(* CODESYS project snapshot.xml
   cds-daemon-config: {"poll_ms": 60, "deny": []}
   cts-project-id: 374e2afd-b7d6-4447-8bd8-ce8e480d827d
   cds-sync-pc: WIN-CODESYS
   cds-sync-folder: ..

Project tree, tasks and I/O mapping:
  PLC_Stabur : PLC Stabur, PSV Electric, order no. psve.ru, version 3.5.16.40
    application Application
      libraries: SysTimeCore, * (System); CmpLog, * (System); CmpErrors, * (System); CmpApp, * (System); Standard, 3.5.22.0 (System); Component Manager, * (System); CmpIecTask, * (System)
      task VISU_TASK (cyclic, interval 100 ms, priority 31) calls VisuElems.Visu_Prg
      task Task (cyclic, interval 200 ms, priority 1) calls MAIN
      data type ST_Bits8
      data type ST_Packed
      function block FB_Logger [ST]: LogADDLong, LogSafe, LogADD, Fmt100
      data type U_Bits8
      program PRG_BitBench [ST]
      visualisation Visualization
      global variables LogComponent
      program MAIN [ST]
      function block FB_BenchRun [ST]
      data type ST_Bools8
      global variables GVL_Bench
      data type U_ExtBits
      data type ST_Bits8Ext
      data type E_BenchMode
      function block FB_Motor [ST]
      global variables GVL_Motors
      function F_Scale [ST]
      global variables GVL_Fixture
      function block FB_Valve [ST]: P_Open, A_Reset, M_Toggle
      LiveTmpFolder/
        global variables GVL_LiveTmp
      interface I_LiveTmp: M_LiveTmp
    Retain_ : Retain, PSV Electric, order no. --0--, version 3.5.16.40
        unmapped channels: Record counter, RETAIN status code, Write
    Leds : Leds, PSV Electro, order no. --0--, version 3.5.16.40
        unmapped channels: LEDs, Screen brightness, Buzzer
  text list GlobalTextList
*)

// PLC_Stabur/Application/ST_Bits8
TYPE ST_Bits8 :
STRUCT
	bit0 : BIT;
	bit1 : BIT;
	bit2 : BIT;
	bit3 : BIT;
	bit4 : BIT;
	bit5 : BIT;
	bit6 : BIT;
	bit7 : BIT;
END_STRUCT
END_TYPE

// PLC_Stabur/Application/ST_Packed
{attribute 'pack_mode' := '0'}
TYPE ST_Packed :
STRUCT
	bTag : BOOL;
	wData : WORD;
END_STRUCT
END_TYPE

// PLC_Stabur/Application/U_Bits8
TYPE U_Bits8 :
UNION
	b : BYTE;
	bits : ST_Bits8;
END_UNION
END_TYPE

// PLC_Stabur/Application/ST_Bools8
TYPE ST_Bools8 :
STRUCT
	b0 : BOOL;
	b1 : BOOL;
	b2 : BOOL;
	b3 : BOOL;
	b4 : BOOL;
	b5 : BOOL;
	b6 : BOOL;
	b7 : BOOL;
END_STRUCT
END_TYPE

// PLC_Stabur/Application/U_ExtBits
TYPE U_ExtBits :
UNION
	b : BYTE;
	bits : ST_Bits8Ext;
END_UNION
END_TYPE

// PLC_Stabur/Application/ST_Bits8Ext
TYPE ST_Bits8Ext EXTENDS ST_Bits8 :
STRUCT
END_STRUCT
END_TYPE

// PLC_Stabur/Application/E_BenchMode
{attribute 'qualified_only'}
TYPE E_BenchMode :
(
	Idle := 0,
	Run := 1,
	Fault := 7
) INT;
END_TYPE

// PLC_Stabur/Application/LogComponent
{attribute 'qualified_only'}
{attribute 'symbol' := 'none'}
VAR_GLOBAL
	BITBENCH : STRING := 'BitBench';	// component name in the runtime log
	sNumFmt  : STRING(80);				// FB_Logger.Fmt100 puts the formatted number here

	logger : FB_Logger;					// the logger itself (production sample)
END_VAR

// PLC_Stabur/Application/GVL_Bench
{attribute 'qualified_only'}
VAR_GLOBAL
	// --- control (written by the host; a run starts itself 50 cycles after start) ---
	xRun			: BOOL;			// rising edge: run the tests again
	xRunUnaligned	: BOOL;			// TRUE: also run B8 (unaligned WORD, may crash)
	sCpuMode		: STRING(40);	// CPU frequency mode, written by the host before a run; printed in the log
	// --- observation ---
	xDone			: BOOL;			// run finished
	nState			: INT;			// state of the PRG_BitBench machine
	nTestIdx		: INT;			// current test 0..21 (a round = one test in one cycle)
	nMeasIdx		: INT;			// how many pairs went into the statistics of the last round
	nIter			: UDINT;		// iterations in one half of a pair (both halves are identical)
	nHeartbeat		: UDINT;		// ++ on every call of the task
	nLastNs			: ULINT;		// duration of the last round (without calibration), ns
	dwSink			: DWORD;		// read sink
	dwSinkW			: DWORD;		// write sink (write baseline)
	// --- results: index 0..10 = B0..B7c, B8 ---
	// Difference = variant - base within a pair, the unit is HUNDREDTHS of ns/operation.
	// The median and the percentiles are computed over the pair differences of one round (NPAIRS = 101).
	medDiffRead		: ARRAY [0..10] OF DINT;	// median of the difference, read
	p25DiffRead		: ARRAY [0..10] OF DINT;	// 25th percentile of the difference
	p75DiffRead		: ARRAY [0..10] OF DINT;	// 75th percentile of the difference
	minDiffRead		: ARRAY [0..10] OF DINT;	// the smallest difference (extreme point)
	minVarRead		: ARRAY [0..10] OF DWORD;	// absolute minimum of the variant, hundredths of ns/op
	minBaseRead		: ARRAY [0..10] OF DWORD;	// absolute minimum of the base, hundredths of ns/op
	nIterRead		: ARRAY [0..10] OF UDINT;	// nIter at the end of the test
	nRoundUsRead	: ARRAY [0..10] OF UDINT;	// duration of the round, us
	medDiffWrite	: ARRAY [0..10] OF DINT;	// median of the difference, write
	p25DiffWrite	: ARRAY [0..10] OF DINT;
	p75DiffWrite	: ARRAY [0..10] OF DINT;
	minDiffWrite	: ARRAY [0..10] OF DINT;
	minVarWrite		: ARRAY [0..10] OF DWORD;
	minBaseWrite	: ARRAY [0..10] OF DWORD;
	nIterWrite		: ARRAY [0..10] OF UDINT;
	nRoundUsWrite	: ARRAY [0..10] OF UDINT;
	nMeasDone		: ARRAY [0..10] OF INT;		// how many pairs went into the result (0 = SKIPPED)
	// --- one-off values ---
	aSizeof			: ARRAY [0..5] OF INT;		// SIZEOF of the types
	// --- enum live check ---
	eMode : E_BenchMode := E_BenchMode.Idle;
	aMode : ARRAY [0..2] OF E_BenchMode := [E_BenchMode.Idle, E_BenchMode.Run, E_BenchMode.Fault];
	// --- test data ---
	stBools			: ST_Bools8;
	stBits			: ST_Bits8;
	uBits			: U_Bits8;
	uExt			: U_ExtBits;
	wData			: WORD;
	dwDataB6		: DWORD;
	stPacked		: ST_Packed;
END_VAR

// PLC_Stabur/Application/GVL_Motors
{attribute 'qualified_only'}
VAR_GLOBAL
	xM1Start : BOOL;
	xM1Stop : BOOL;
	xM1Feedback : BOOL;
	xM1Reset : BOOL;
	xM1Run : BOOL;
	xM1Fault : BOOL;
	nM1Starts : UDINT;
	fbMotor1 : FB_Motor;

	xM2Start : BOOL;
	xM2Stop : BOOL;
	xM2Feedback : BOOL;
	xM2Reset : BOOL;
	xM2Run : BOOL;
	xM2Fault : BOOL;
	nM2Starts : UDINT;
	fbMotor2 : FB_Motor;
END_VAR

// PLC_Stabur/Application/GVL_Fixture
VAR_GLOBAL
	rScaled : REAL;
	xValveOpen : BOOL;
	fbValve : FB_Valve;
	nTicks : UDINT;
END_VAR

// PLC_Stabur/Application/LiveTmpFolder/GVL_LiveTmp
VAR_GLOBAL
	xLiveTmp : BOOL;
END_VAR

// PLC_Stabur/Application/MAIN
PROGRAM MAIN
(* t76 timing probe *)
VAR
	eObservedMode : E_BenchMode;
END_VAR

// Self-contained bit-access benchmark: it starts itself 50 cycles after the
// application starts, writes its report to the runtime log, and repeats on GVL_Bench.xRun.
// Project created with the cds-text-sync daemon and LLM agent.
PRG_BitBench();
eObservedMode := GVL_Bench.eMode;

GVL_Motors.fbMotor1(
	xStart := GVL_Motors.xM1Start,
	xStop := GVL_Motors.xM1Stop,
	xFeedback := GVL_Motors.xM1Feedback,
	xReset := GVL_Motors.xM1Reset,
	xRun => GVL_Motors.xM1Run,
	xFault => GVL_Motors.xM1Fault,
	nStarts => GVL_Motors.nM1Starts);
GVL_Motors.fbMotor2(
	xStart := GVL_Motors.xM2Start,
	xStop := GVL_Motors.xM2Stop,
	xFeedback := GVL_Motors.xM2Feedback,
	xReset := GVL_Motors.xM2Reset,
	xRun => GVL_Motors.xM2Run,
	xFault => GVL_Motors.xM2Fault,
	nStarts => GVL_Motors.nM2Starts);

// Fixture: exercise the function, property, action and interface kinds.
GVL_Fixture.nTicks := GVL_Fixture.nTicks + 1;
GVL_Fixture.rScaled := F_Scale(UDINT_TO_REAL(GVL_Fixture.nTicks), 0.5);
IF GVL_Fixture.nTicks MOD 10 = 0 THEN
	GVL_Fixture.fbValve.M_Toggle();
END_IF
GVL_Fixture.xValveOpen := GVL_Fixture.fbValve.P_Open;

END_PROGRAM

// PLC_Stabur/Application/PRG_BitBench
(*
BitBench — a self-contained benchmark of the cost of bit access.

Project created with the cds-text-sync daemon and LLM agent.
Bench: PLC_Stabur (RK3568, 4x ARM Cortex-A55), CODESYS Control 3.5.16.40,
task t#200 ms, timer SysTimeGetNs on the PLC.

RUN ORDER (counted in task cycles):
  PLC on / application started
  -> wait START_WAIT cycles (50 = 10 s)
  -> round 1: one test ENTIRELY in one cycle
  -> wait GAP_WAIT cycles (5 = 1 s)
  -> round 2 ... and so on up to the last test
  -> conclusion (Conclusion) and 'BitBench: done'.
The 20 tests (B0..B7c read and write) take about 30 s; B8 takes two more rounds.

THE METHOD OF ONE ROUND - PAIRED MEASUREMENTS.
The calibration (CAL_N iterations) chooses nIter so that one half of a pair runs
for about TARGET_EACH_NS. Then WARM_PAIRS warm-up pairs and NPAIRS measured pairs
in a row: a pair is the baseline and the variant with the same nIter, the order
alternates (even pair base -> variant, odd pair the other way round). The result
of a pair is the difference (variant - base) in hundredths of ns/operation. The
differences are sorted at the end of the round; Result is the median, with p25,
p75 and min beside it.

A round is limited by ROUND_BUDGET_NS: if the pairs did not fit, the round is cut
short and is computed from the pairs that made it (fewer than MIN_PAIRS -
SKIPPED). We reset the statistics of the task (CmpIecTask) in the last cycle of
the pause before the round and read them in the first cycle after it: the cycle
max is the round itself.

Restart. A run starts over (from the START_WAIT pause) if:
  - the application was downloaded or reset (the variables are initialised);
  - more than RESTART_GAP_NS passed between two cycles (Online -> Stop/Start:
    the variables survive, but the task was stopped);
  - a rising edge on GVL_Bench.xRun (then the pause is GAP_WAIT, not START_WAIT).
B8 (an unaligned WORD in a STRUCT with pack_mode 0) runs only when
GVL_Bench.xRunUnaligned is set, because it may raise an exception.

We keep the log strings no longer than 120 characters (the runtime cuts a record
at 127); anything longer is sent by LogSafe in pieces.
*)

PROGRAM PRG_BitBench
VAR CONSTANT
	// --- schedule, in task cycles ---
	START_WAIT	: INT := 50;			// after the application starts
	GAP_WAIT	: INT := 5;				// between rounds
	TASK_NS		: ULINT := 200000000;	// task period, ns (t#200 ms)
	RESTART_GAP_NS : ULINT := 1000000000;	// a gap between cycles longer than 1 s = the task was stopped
	// --- method ---
	CAL_N		: UDINT := 1000;		// iterations in the calibration half
	WARM_PAIRS	: INT := 5;				// warm-up pairs (they do not enter the statistics)
	NPAIRS		: INT := 101;			// measured pairs per test (odd - the median is unambiguous)
	MIN_PAIRS	: INT := 21;			// fewer - the test is SKIPPED
	MIN_ITER	: UDINT := 50;
	MAX_ITER	: UDINT := 2000000;
	TARGET_EACH_NS : ULINT := 200000;	// target duration of half a pair, ns (0.2 ms)
	ROUND_BUDGET_NS : ULINT := 80000000;	// round limit, ns (80 ms = 40 % of the cycle)
	// --- tests ---
	IDX_LAST_MAIN : INT := 19;			// 0..9 read B0..B7c, 10..19 write
	IDX_LAST	: INT := 21;			// 20 = read B8, 21 = write B8
	// --- states ---
	ST_IDLE		: INT := 0;				// no run in progress
	ST_WAIT		: INT := 10;			// pause before a round (nWait cycles)
	ST_ROUND	: INT := 20;			// round: one test in this cycle
	ST_DONE		: INT := 100;			// run finished
END_VAR
VAR
	// --- start and restart ---
	xInit		: BOOL;			// FALSE after a download/reset: the first cycle
	xRunPrev	: BOOL;
	tNow		: ULINT;
	tPrevCycle	: ULINT;
	// --- state machine ---
	nFsm		: INT;
	nWait		: INT;			// how many cycles of the pause are left
	xHeadDone	: BOOL;			// the run header has already been printed
	xStatPending : BOOL;		// print the statistics of the task for the round in this cycle
	nTestNo		: INT;			// 0..21
	// --- current test ---
	nMode		: INT;			// 0 = read, 1 = write
	nVariant	: INT;			// 0..10
	nIterCur	: UDINT;		// nIter of the round: the same for both halves of every pair
	// --- statistics of the task itself (CmpIecTask, as in FB_TaskInfo from a production sample) ---
	pTaskInfo	: POINTER TO Task_Info2;
	resTask		: UDINT;
	// --- measurements ---
	fbRun		: FB_BenchRun;
	tBase		: ULINT;
	tVar		: ULINT;
	tPair		: ULINT;
	tRound0		: ULINT;
	tRoundNs	: ULINT;		// duration of the round (without calibration), ns
	uCalBase	: ULINT;
	uCalVar		: ULINT;
	aDiff		: ARRAY [0..100] OF DINT;	// pair differences (NPAIRS = 101)
	nMeasCnt	: INT;
	xCut		: BOOL;			// the round was cut by ROUND_BUDGET_NS
	uMaxPair	: ULINT;
	uMinVar		: ULINT;		// absolute minimum of the variant, hundredths of ns/op
	uMinBase	: ULINT;
	dNew		: DINT;
	dMed		: DINT;
	dP25		: DINT;
	dP75		: DINT;
	dMn			: DINT;
	// --- processing ---
	p			: INT;
	i			: INT;
	j			: INT;
	uTmp		: ULINT;
	dwRes		: DWORD;
	xTimerBad	: BOOL;
	dRead		: DINT;
	dWrite		: DINT;
	dWorst		: DINT;
	dTmp		: DINT;
	// --- strings ---
	sMsg		: STRING(255);
	sName		: STRING(40);
	sWhat		: STRING(80);
END_VAR

// ===================== 1. start, restart, manual run =====================
dwRes := SysTimeGetNs(tNow);

IF NOT xInit THEN
	// the first cycle after a download or a reset
	xInit := TRUE;
	nFsm := ST_WAIT;
	nWait := START_WAIT;
	xHeadDone := FALSE;
	xStatPending := FALSE;
	LogComponent.logger.LogSafe(LogComponent.BITBENCH, CmpLog.LogClass.LOG_INFO,
		'BitBench: application started, first round after 50 cycles');
ELSIF tPrevCycle <> 0 AND tNow - tPrevCycle > RESTART_GAP_NS THEN
	// the task was stopped (Online -> Stop/Start): we start the run over
	nFsm := ST_WAIT;
	nWait := START_WAIT;
	xHeadDone := FALSE;
	xStatPending := FALSE;
	LogComponent.logger.LogSafe(LogComponent.BITBENCH, CmpLog.LogClass.LOG_INFO,
		'BitBench: restart after a stop, first round after 50 cycles');
END_IF
tPrevCycle := tNow;

IF GVL_Bench.xRun AND NOT xRunPrev THEN
	nFsm := ST_WAIT;
	nWait := GAP_WAIT;
	xHeadDone := FALSE;
	xStatPending := FALSE;
END_IF
xRunPrev := GVL_Bench.xRun;

// ===================== 2. task statistics for the previous round =====================
IF xStatPending THEN
	xStatPending := FALSE;
	IF pTaskInfo <> 0 THEN
		sMsg := CONCAT('Task      ', sName);
		sMsg := CONCAT(sMsg, ': cycle max ');
		sMsg := CONCAT(sMsg, DWORD_TO_STRING(pTaskInfo^.dwMaxCycleTime));
		sMsg := CONCAT(sMsg, ' us, jitter max ');
		sMsg := CONCAT(sMsg, DINT_TO_STRING(pTaskInfo^.iJitterMax));
		sMsg := CONCAT(sMsg, ' us, min ');
		sMsg := CONCAT(sMsg, DINT_TO_STRING(pTaskInfo^.iJitterMin));
		sMsg := CONCAT(sMsg, ' us');
		LogComponent.logger.LogSafe(LogComponent.BITBENCH, CmpLog.LogClass.LOG_INFO, sMsg);
	END_IF
END_IF

// ===================== 3. state machine =====================
CASE nFsm OF
ST_IDLE:
	;	// waiting for xRun or a restart

ST_WAIT:	// pause; the last cycle of the pause prepares the round
	nWait := nWait - 1;
	IF nWait <= 0 THEN
		IF NOT xHeadDone THEN
			xHeadDone := TRUE;
			nTestNo := 0;
			xTimerBad := FALSE;
			GVL_Bench.xDone := FALSE;
			GVL_Bench.dwSink := 0;
			GVL_Bench.dwSinkW := 0;
			// clear the results of the previous run: after a SKIPPED or a crash
			// the GVL must not keep numbers from the previous run
			FOR i := 0 TO 10 DO
				GVL_Bench.medDiffRead[i] := 0;
				GVL_Bench.p25DiffRead[i] := 0;
				GVL_Bench.p75DiffRead[i] := 0;
				GVL_Bench.minDiffRead[i] := 0;
				GVL_Bench.minVarRead[i] := 0;
				GVL_Bench.minBaseRead[i] := 0;
				GVL_Bench.nIterRead[i] := 0;
				GVL_Bench.nRoundUsRead[i] := 0;
				GVL_Bench.medDiffWrite[i] := 0;
				GVL_Bench.p25DiffWrite[i] := 0;
				GVL_Bench.p75DiffWrite[i] := 0;
				GVL_Bench.minDiffWrite[i] := 0;
				GVL_Bench.minVarWrite[i] := 0;
				GVL_Bench.minBaseWrite[i] := 0;
				GVL_Bench.nIterWrite[i] := 0;
				GVL_Bench.nRoundUsWrite[i] := 0;
				GVL_Bench.nMeasDone[i] := 0;
			END_FOR
			GVL_Bench.nIter := 0;
			GVL_Bench.nLastNs := 0;
			GVL_Bench.nMeasIdx := 0;

			// the run header
			LogComponent.logger.LogSafe(LogComponent.BITBENCH, CmpLog.LogClass.LOG_INFO,
				'BitBench: project created with cds-text-sync daemon and LLM agent');

			sMsg := CONCAT('BitBench: start, CPU mode ', GVL_Bench.sCpuMode);
			LogComponent.logger.LogSafe(LogComponent.BITBENCH, CmpLog.LogClass.LOG_INFO, sMsg);

			sMsg := 'BitBench: CPU RK3568 4x ARM Cortex-A55, task t#';
			sMsg := CONCAT(sMsg, ULINT_TO_STRING(TASK_NS / 1000000));
			sMsg := CONCAT(sMsg, ' ms, timer SysTimeGetNs on the PLC');
			LogComponent.logger.LogSafe(LogComponent.BITBENCH, CmpLog.LogClass.LOG_INFO, sMsg);

			sMsg := 'BitBench: 1 round = 1 test in one cycle, ';
			sMsg := CONCAT(sMsg, INT_TO_STRING(GAP_WAIT));
			sMsg := CONCAT(sMsg, ' cycles between rounds, round limit ');
			sMsg := CONCAT(sMsg, ULINT_TO_STRING(ROUND_BUDGET_NS / 1000000));
			sMsg := CONCAT(sMsg, ' ms');
			LogComponent.logger.LogSafe(LogComponent.BITBENCH, CmpLog.LogClass.LOG_INFO, sMsg);

			sMsg := 'BitBench: round = ';
			sMsg := CONCAT(sMsg, INT_TO_STRING(WARM_PAIRS));
			sMsg := CONCAT(sMsg, ' warm-up + ');
			sMsg := CONCAT(sMsg, INT_TO_STRING(NPAIRS));
			sMsg := CONCAT(sMsg, ' measured pairs (base and variant, same nIter), half ~');
			LogComponent.logger.Fmt100(ULINT_TO_DINT(TARGET_EACH_NS / 10000), FALSE);
			sMsg := CONCAT(sMsg, LogComponent.sNumFmt);
			sMsg := CONCAT(sMsg, ' ms');
			LogComponent.logger.LogSafe(LogComponent.BITBENCH, CmpLog.LogClass.LOG_INFO, sMsg);

			GVL_Bench.aSizeof[0] := SIZEOF(GVL_Bench.stBools);
			GVL_Bench.aSizeof[1] := SIZEOF(GVL_Bench.stBits);
			GVL_Bench.aSizeof[2] := SIZEOF(GVL_Bench.uBits);
			GVL_Bench.aSizeof[3] := SIZEOF(GVL_Bench.uExt);
			GVL_Bench.aSizeof[4] := SIZEOF(GVL_Bench.stPacked);
			GVL_Bench.aSizeof[5] := SIZEOF(GVL_Bench.wData);

			sMsg := 'Memory: 8 BOOL in a STRUCT = ';
			sMsg := CONCAT(sMsg, INT_TO_STRING(GVL_Bench.aSizeof[0]));
			sMsg := CONCAT(sMsg, ' B, 8 BIT in a STRUCT = ');
			sMsg := CONCAT(sMsg, INT_TO_STRING(GVL_Bench.aSizeof[1]));
			sMsg := CONCAT(sMsg, ' B, UNION of 8 BIT = ');
			sMsg := CONCAT(sMsg, INT_TO_STRING(GVL_Bench.aSizeof[2]));
			sMsg := CONCAT(sMsg, ' B');
			LogComponent.logger.LogSafe(LogComponent.BITBENCH, CmpLog.LogClass.LOG_INFO, sMsg);

			sMsg := 'Memory: the same UNION + EXTENDS = ';
			sMsg := CONCAT(sMsg, INT_TO_STRING(GVL_Bench.aSizeof[3]));
			sMsg := CONCAT(sMsg, ' B, WORD = ');
			sMsg := CONCAT(sMsg, INT_TO_STRING(GVL_Bench.aSizeof[5]));
			sMsg := CONCAT(sMsg, ' B, pack_mode 0 (WORD after BOOL) = ');
			sMsg := CONCAT(sMsg, INT_TO_STRING(GVL_Bench.aSizeof[4]));
			sMsg := CONCAT(sMsg, ' B');
			LogComponent.logger.LogSafe(LogComponent.BITBENCH, CmpLog.LogClass.LOG_INFO, sMsg);

			LogComponent.logger.LogSafe(LogComponent.BITBENCH, CmpLog.LogClass.LOG_INFO,
				'Base  read: dwSink := dwSink + 1; write: dwSinkW := UDINT_TO_DWORD(k AND 1)');

			IF pTaskInfo = 0 THEN
				pTaskInfo := IecTaskGetInfo3(hIecTask := IecTaskGetCurrent(ADR(resTask)),
				                             pResult := ADR(resTask));
			END_IF
		END_IF

		// the task statistics from this moment on are the statistics of the round
		IecTaskResetStatistics(IecTaskGetCurrent(ADR(resTask)));
		nFsm := ST_ROUND;
	END_IF

ST_ROUND:	// one test entirely in this cycle
	// ---------- which test ----------
	IF nTestNo < 10 THEN
		nMode := 0;
		nVariant := nTestNo;
	ELSIF nTestNo <= IDX_LAST_MAIN THEN
		nMode := 1;
		nVariant := nTestNo - 10;
	ELSIF nTestNo = IDX_LAST_MAIN + 1 THEN
		nMode := 0;
		nVariant := 10;
	ELSE
		nMode := 1;
		nVariant := 10;
	END_IF

	CASE nVariant OF
	0:	sName := 'B0 empty loop';
		sWhat := 'control: the variant is the base itself, expect 0';
	1:	sName := 'B1 BOOL fields';
		sWhat := '8 BOOL in a STRUCT, 1 byte each - the reference for the bit tests';
	2:	sName := 'B2 BIT fields';
		sWhat := '8 BIT packed into 1 byte - the write is a read-modify-write';
	3:	sName := 'B3 UNION+EXTENDS';
		sWhat := 'bit via a UNION that EXTENDS ST_Bits8; watch C0542';
	4:	sName := 'B4 UNION';
		sWhat := 'the same 8 BIT in a UNION, without EXTENDS';
	5:	sName := 'B5 WORD.3';
		sWhat := 'bit access to a WORD by dot: wData.3, 16 bits in 2 B';
	6:	sName := 'B6 mask var index';
		sWhat := 'mask (SHR(dwData, i) AND 1), no bit instruction';
	7:	sName := 'B7a 8 BOOL';
		sWhat := '8 BOOL one by one - one iteration = 8 accesses';
	8:	sName := 'B7b byte';
		sWhat := 'all 8 bits as one BYTE - one iteration = 1 access';
	9:	sName := 'B7c word';
		sWhat := 'all 16 bits as one WORD - one iteration = 1 access';
	10:	sName := 'B8 unaligned WORD';
		sWhat := 'pack_mode 0, wData.3 unaligned - the test may raise an exception';
	ELSE
		sName := 'B? unknown';
		sWhat := 'unknown variant';
	END_CASE

	sMsg := CONCAT('Testing ', sName);
	IF nMode = 0 THEN
		sMsg := CONCAT(sMsg, ' (read): ');
	ELSE
		sMsg := CONCAT(sMsg, ' (write): ');
	END_IF
	sMsg := CONCAT(sMsg, sWhat);
	LogComponent.logger.LogSafe(LogComponent.BITBENCH, CmpLog.LogClass.LOG_INFO, sMsg);

	IF nVariant = 10 THEN
		LogComponent.logger.LogSafe(LogComponent.BITBENCH, CmpLog.LogClass.LOG_WARNING,
			'B8 warning: unaligned WORD in a STRUCT with pack_mode 0; an exception here means the app restarts');
	END_IF

	// ---------- calibration: nIter for TARGET_EACH_NS from the slower half ----------
	fbRun(nWhich := 0, nMode := nMode, nVariant := nVariant, nIter := CAL_N);
	uCalBase := fbRun.tDur;
	IF fbRun.dwRes <> 0 THEN
		dwRes := fbRun.dwRes;
	END_IF
	fbRun(nWhich := 1, nMode := nMode, nVariant := nVariant, nIter := CAL_N);
	uCalVar := fbRun.tDur;
	IF fbRun.dwRes <> 0 THEN
		dwRes := fbRun.dwRes;
	END_IF

	uTmp := uCalBase;
	IF uCalVar > uTmp THEN
		uTmp := uCalVar;
	END_IF
	IF uTmp <> 0 THEN
		uTmp := (TARGET_EACH_NS * CAL_N) / uTmp;
	ELSE
		uTmp := MIN_ITER;
	END_IF
	IF uTmp < MIN_ITER THEN
		uTmp := MIN_ITER;
	END_IF
	IF uTmp > MAX_ITER THEN
		uTmp := MAX_ITER;
	END_IF
	nIterCur := ULINT_TO_UDINT(uTmp);
	GVL_Bench.nIter := nIterCur;

	// ---------- pairs: warm-up, then measured ----------
	nMeasCnt := 0;
	xCut := FALSE;
	uMaxPair := 0;
	uMinVar := 16#FFFFFFFFFFFFFFFF;
	uMinBase := 16#FFFFFFFFFFFFFFFF;
	SysTimeGetNs(tRound0);

	FOR p := 0 TO WARM_PAIRS + NPAIRS - 1 DO
		IF (p MOD 2) = 0 THEN
			fbRun(nWhich := 0, nMode := nMode, nVariant := nVariant, nIter := nIterCur);
			tBase := fbRun.tDur;
			fbRun(nWhich := 1, nMode := nMode, nVariant := nVariant, nIter := nIterCur);
			tVar := fbRun.tDur;
		ELSE
			fbRun(nWhich := 1, nMode := nMode, nVariant := nVariant, nIter := nIterCur);
			tVar := fbRun.tDur;
			fbRun(nWhich := 0, nMode := nMode, nVariant := nVariant, nIter := nIterCur);
			tBase := fbRun.tDur;
		END_IF
		IF fbRun.dwRes <> 0 THEN
			dwRes := fbRun.dwRes;
		END_IF

		IF p >= WARM_PAIRS THEN
			tPair := tBase + tVar;
			IF tPair > uMaxPair THEN
				uMaxPair := tPair;
			END_IF
			// the difference in hundredths of ns/op: each half is normalised separately
			uTmp := (tVar * 100) / nIterCur;
			IF uTmp < uMinVar THEN
				uMinVar := uTmp;
			END_IF
			dNew := ULINT_TO_DINT(uTmp);
			uTmp := (tBase * 100) / nIterCur;
			IF uTmp < uMinBase THEN
				uMinBase := uTmp;
			END_IF
			dNew := dNew - ULINT_TO_DINT(uTmp);
			aDiff[nMeasCnt] := dNew;
			nMeasCnt := nMeasCnt + 1;
		END_IF

		// round limit: the task cycle must not overrun the budget
		SysTimeGetNs(tPair);
		IF tPair - tRound0 > ROUND_BUDGET_NS THEN
			xCut := TRUE;
			EXIT;
		END_IF
	END_FOR

	SysTimeGetNs(tPair);
	tRoundNs := tPair - tRound0;
	GVL_Bench.nLastNs := tRoundNs;
	GVL_Bench.nMeasIdx := nMeasCnt;

	// ---------- insertion sort (101 elements, once per round) ----------
	FOR i := 1 TO nMeasCnt - 1 DO
		dNew := aDiff[i];
		j := i - 1;
		WHILE j >= 0 DO
			IF aDiff[j] > dNew THEN
				aDiff[j + 1] := aDiff[j];
				j := j - 1;
			ELSE
				EXIT;
			END_IF
		END_WHILE
		aDiff[j + 1] := dNew;
	END_FOR

	// ---------- round result ----------
	sMsg := CONCAT('Result  ', sName);
	IF nMode = 0 THEN
		sMsg := CONCAT(sMsg, ' (read): ');
	ELSE
		sMsg := CONCAT(sMsg, ' (write): ');
	END_IF

	IF nMeasCnt >= MIN_PAIRS THEN
		dMn := aDiff[0];
		dP25 := aDiff[nMeasCnt / 4];
		dMed := aDiff[nMeasCnt / 2];
		dP75 := aDiff[(nMeasCnt * 3) / 4];

		IF nMode = 0 THEN
			GVL_Bench.medDiffRead[nVariant] := dMed;
			GVL_Bench.p25DiffRead[nVariant] := dP25;
			GVL_Bench.p75DiffRead[nVariant] := dP75;
			GVL_Bench.minDiffRead[nVariant] := dMn;
			GVL_Bench.minVarRead[nVariant] := ULINT_TO_DWORD(uMinVar);
			GVL_Bench.minBaseRead[nVariant] := ULINT_TO_DWORD(uMinBase);
			GVL_Bench.nIterRead[nVariant] := nIterCur;
			GVL_Bench.nRoundUsRead[nVariant] := ULINT_TO_UDINT(tRoundNs / 1000);
		ELSE
			GVL_Bench.medDiffWrite[nVariant] := dMed;
			GVL_Bench.p25DiffWrite[nVariant] := dP25;
			GVL_Bench.p75DiffWrite[nVariant] := dP75;
			GVL_Bench.minDiffWrite[nVariant] := dMn;
			GVL_Bench.minVarWrite[nVariant] := ULINT_TO_DWORD(uMinVar);
			GVL_Bench.minBaseWrite[nVariant] := ULINT_TO_DWORD(uMinBase);
			GVL_Bench.nIterWrite[nVariant] := nIterCur;
			GVL_Bench.nRoundUsWrite[nVariant] := ULINT_TO_UDINT(tRoundNs / 1000);
		END_IF
		GVL_Bench.nMeasDone[nVariant] := nMeasCnt;

		// Result - the median of the pair differences, the sign comes from the number itself
		LogComponent.logger.Fmt100(dMed, TRUE);
		sMsg := CONCAT(sMsg, LogComponent.sNumFmt);
		sMsg := CONCAT(sMsg, ' ns/op vs base (');
		sMsg := CONCAT(sMsg, INT_TO_STRING(nMeasCnt));
		sMsg := CONCAT(sMsg, ': p25 ');
		LogComponent.logger.Fmt100(dP25, TRUE);
		sMsg := CONCAT(sMsg, LogComponent.sNumFmt);
		sMsg := CONCAT(sMsg, ', p75 ');
		LogComponent.logger.Fmt100(dP75, TRUE);
		sMsg := CONCAT(sMsg, LogComponent.sNumFmt);
		sMsg := CONCAT(sMsg, ', min ');
		LogComponent.logger.Fmt100(dMn, TRUE);
		sMsg := CONCAT(sMsg, LogComponent.sNumFmt);
		sMsg := CONCAT(sMsg, '), nIter ');
		sMsg := CONCAT(sMsg, UDINT_TO_STRING(nIterCur));
		LogComponent.logger.LogSafe(LogComponent.BITBENCH, CmpLog.LogClass.LOG_INFO, sMsg);
	ELSE
		// SKIPPED - explicitly, and nothing is left in the GVL
		IF nMode = 0 THEN
			GVL_Bench.medDiffRead[nVariant] := 0;
		ELSE
			GVL_Bench.medDiffWrite[nVariant] := 0;
		END_IF
		GVL_Bench.nMeasDone[nVariant] := 0;
		sMsg := CONCAT(sMsg, 'SKIPPED, only ');
		sMsg := CONCAT(sMsg, INT_TO_STRING(nMeasCnt));
		sMsg := CONCAT(sMsg, ' pairs fit the round limit');
		LogComponent.logger.LogSafe(LogComponent.BITBENCH, CmpLog.LogClass.LOG_ERROR, sMsg);
	END_IF

	// Round - the duration of the round and the absolute minima of both halves
	sMsg := CONCAT('Round     ', sName);
	sMsg := CONCAT(sMsg, ': ');
	LogComponent.logger.Fmt100(ULINT_TO_DINT(tRoundNs / 10000), FALSE);
	sMsg := CONCAT(sMsg, LogComponent.sNumFmt);
	sMsg := CONCAT(sMsg, ' ms');
	IF xCut THEN
		sMsg := CONCAT(sMsg, ' (cut at the limit)');
	END_IF
	sMsg := CONCAT(sMsg, ', max pair ');
	LogComponent.logger.Fmt100(ULINT_TO_DINT(uMaxPair / 10000), FALSE);
	sMsg := CONCAT(sMsg, LogComponent.sNumFmt);
	sMsg := CONCAT(sMsg, ' ms, min var ');
	LogComponent.logger.Fmt100(ULINT_TO_DINT(uMinVar), FALSE);
	sMsg := CONCAT(sMsg, LogComponent.sNumFmt);
	sMsg := CONCAT(sMsg, ' / base ');
	LogComponent.logger.Fmt100(ULINT_TO_DINT(uMinBase), FALSE);
	sMsg := CONCAT(sMsg, LogComponent.sNumFmt);
	sMsg := CONCAT(sMsg, ' ns/op');
	LogComponent.logger.LogSafe(LogComponent.BITBENCH, CmpLog.LogClass.LOG_INFO, sMsg);

	// ---------- next round, conclusion, or the end ----------
	xStatPending := TRUE;
	nTestNo := nTestNo + 1;

	IF nTestNo = IDX_LAST_MAIN + 1 THEN
		// Conclusion from the MEDIANS of the pair differences; min beside it
		dRead := GVL_Bench.medDiffRead[2] - GVL_Bench.medDiffRead[1];
		dWrite := GVL_Bench.medDiffWrite[2] - GVL_Bench.medDiffWrite[1];

		LogComponent.logger.LogSafe(LogComponent.BITBENCH, CmpLog.LogClass.LOG_INFO, '=========');

		sMsg := 'Conclusion: BIT vs BOOL fields (B2 - B1), median read ';
		LogComponent.logger.Fmt100(dRead, TRUE);
		sMsg := CONCAT(sMsg, LogComponent.sNumFmt);
		sMsg := CONCAT(sMsg, ' (min ');
		LogComponent.logger.Fmt100(GVL_Bench.minDiffRead[2] - GVL_Bench.minDiffRead[1], TRUE);
		sMsg := CONCAT(sMsg, LogComponent.sNumFmt);
		sMsg := CONCAT(sMsg, '), write ');
		LogComponent.logger.Fmt100(dWrite, TRUE);
		sMsg := CONCAT(sMsg, LogComponent.sNumFmt);
		sMsg := CONCAT(sMsg, ' (min ');
		LogComponent.logger.Fmt100(GVL_Bench.minDiffWrite[2] - GVL_Bench.minDiffWrite[1], TRUE);
		sMsg := CONCAT(sMsg, LogComponent.sNumFmt);
		sMsg := CONCAT(sMsg, ') ns/op');
		LogComponent.logger.LogSafe(LogComponent.BITBENCH, CmpLog.LogClass.LOG_INFO, sMsg);

		IF dWrite > dRead THEN
			dWorst := dWrite;
		ELSE
			dWorst := dRead;
		END_IF
		IF dWorst < 0 THEN
			dWorst := 0;
		END_IF

		// dWorst is in hundredths of ns/op, so 1000 accesses = dWorst/100 us.
		// The share of the cycle in ppm = dWorst * 10 ns * 1e6 / TASK_NS; printed in hundredths of ppm.
		sMsg := 'Conclusion: 1000 bit accesses cost ';
		LogComponent.logger.Fmt100(dWorst, FALSE);
		sMsg := CONCAT(sMsg, LogComponent.sNumFmt);
		sMsg := CONCAT(sMsg, ' us = ');
		LogComponent.logger.Fmt100(LINT_TO_DINT(DINT_TO_LINT(dWorst) * 1000000000 / ULINT_TO_LINT(TASK_NS)), FALSE);
		sMsg := CONCAT(sMsg, LogComponent.sNumFmt);
		sMsg := CONCAT(sMsg, ' ppm of the ');
		sMsg := CONCAT(sMsg, ULINT_TO_STRING(TASK_NS / 1000000));
		sMsg := CONCAT(sMsg, ' ms task cycle');
		LogComponent.logger.LogSafe(LogComponent.BITBENCH, CmpLog.LogClass.LOG_INFO, sMsg);

		dTmp := GVL_Bench.medDiffRead[7] - GVL_Bench.medDiffRead[8];
		sMsg := 'Conclusion: 8 BOOL one by one vs 1 BYTE read (B7a - B7b), median ';
		LogComponent.logger.Fmt100(dTmp, TRUE);
		sMsg := CONCAT(sMsg, LogComponent.sNumFmt);
		sMsg := CONCAT(sMsg, ' (min ');
		LogComponent.logger.Fmt100(GVL_Bench.minDiffRead[7] - GVL_Bench.minDiffRead[8], TRUE);
		sMsg := CONCAT(sMsg, LogComponent.sNumFmt);
		sMsg := CONCAT(sMsg, ') ns/iteration');
		LogComponent.logger.LogSafe(LogComponent.BITBENCH, CmpLog.LogClass.LOG_INFO, sMsg);

		dTmp := GVL_Bench.medDiffRead[3] - GVL_Bench.medDiffRead[4];
		sMsg := 'Conclusion: UNION+EXTENDS vs UNION (B3 - B4), median read ';
		LogComponent.logger.Fmt100(dTmp, TRUE);
		sMsg := CONCAT(sMsg, LogComponent.sNumFmt);
		sMsg := CONCAT(sMsg, ', write ');
		LogComponent.logger.Fmt100(GVL_Bench.medDiffWrite[3] - GVL_Bench.medDiffWrite[4], TRUE);
		sMsg := CONCAT(sMsg, LogComponent.sNumFmt);
		sMsg := CONCAT(sMsg, ' ns/op');
		LogComponent.logger.LogSafe(LogComponent.BITBENCH, CmpLog.LogClass.LOG_INFO, sMsg);

		IF GVL_Bench.xRunUnaligned THEN
			nWait := GAP_WAIT;
			nFsm := ST_WAIT;
		ELSE
			LogComponent.logger.LogSafe(LogComponent.BITBENCH, CmpLog.LogClass.LOG_INFO,
				'B8 skipped: GVL_Bench.xRunUnaligned = FALSE');
			nFsm := ST_DONE;
		END_IF
	ELSIF nTestNo > IDX_LAST THEN
		nFsm := ST_DONE;
	ELSE
		nWait := GAP_WAIT;
		nFsm := ST_WAIT;
	END_IF

ST_DONE:	// run finished
	GVL_Bench.xDone := TRUE;
	LogComponent.logger.LogSafe(LogComponent.BITBENCH, CmpLog.LogClass.LOG_INFO, 'BitBench: done');
	nFsm := ST_IDLE;

ELSE
	nFsm := ST_IDLE;
END_CASE

// timer return code: 0 = success; non-zero - the measurements are garbage
IF dwRes <> 0 AND NOT xTimerBad THEN
	xTimerBad := TRUE;
	sMsg := CONCAT('SysTimeGetNs error code ', DWORD_TO_STRING(dwRes));
	LogComponent.logger.LogSafe(LogComponent.BITBENCH, CmpLog.LogClass.LOG_ERROR, sMsg);
END_IF

// ===================== 4. observation =====================
GVL_Bench.nState := nFsm;
GVL_Bench.nTestIdx := nTestNo;
GVL_Bench.nHeartbeat := GVL_Bench.nHeartbeat + 1;

END_PROGRAM

// PLC_Stabur/Application/FB_BenchRun
(*
FB_BenchRun — one benchmark loop body: baseline or variant, nIter iterations.

One call = one measured half of a pair. The base and the variant live in the same
block and at the same nesting level, so that the dispatch overhead is the same
and only the loop body differs.

Baseline:
  read - GVL_Bench.dwSink := dwSink + 1 (the same shape as the read variants);
  write - GVL_Bench.dwSinkW := UDINT_TO_DWORD(k AND 1), that is, writing a
  computed value into a separate DWORD sink without touching bits.
The timer is SysTimeGetNs on the PLC (as before, one measurement = one loop pass).

nIter is chosen by the calibration in PRG_BitBench: half of a pair is about
0.2 ms, the whole round (one test) is no more than 80 ms of the t#200 ms cycle.
*)

FUNCTION_BLOCK FB_BenchRun
VAR_INPUT
	nWhich		: INT;			// 0 = baseline, 1 = variant
	nMode		: INT;			// 0 = read, 1 = write
	nVariant	: INT;			// 0..10
	nIter		: UDINT;		// iterations in the loop
END_VAR
VAR_OUTPUT
	tDur		: ULINT;		// duration of the loop, ns
	dwRes		: DWORD;		// return code of SysTimeGetNs (0 = success)
END_VAR
VAR
	k			: UDINT;
	t0			: ULINT;
	t1			: ULINT;
END_VAR

dwRes := SysTimeGetNs(t0);

IF nWhich = 0 THEN
	// ---------------- baseline ----------------
	IF nMode = 0 THEN
		FOR k := 1 TO nIter DO
			GVL_Bench.dwSink := GVL_Bench.dwSink + 1;
		END_FOR
	ELSE
		FOR k := 1 TO nIter DO
			GVL_Bench.dwSinkW := UDINT_TO_DWORD(k AND 1);
		END_FOR
	END_IF
ELSE
	// ---------------- variant ----------------
	IF nMode = 0 THEN		// ---------- READ ----------
		CASE nVariant OF
		0:	// B0 baseline (the same code as the base - a check of the method)
			FOR k := 1 TO nIter DO
				GVL_Bench.dwSink := GVL_Bench.dwSink + 1;
			END_FOR
		1:	// B1 BOOL field of a STRUCT
			FOR k := 1 TO nIter DO
				GVL_Bench.dwSink := GVL_Bench.dwSink + BOOL_TO_DWORD(GVL_Bench.stBools.b3);
			END_FOR
		2:	// B2 BIT field of a STRUCT
			FOR k := 1 TO nIter DO
				GVL_Bench.dwSink := GVL_Bench.dwSink + BOOL_TO_DWORD(GVL_Bench.stBits.bit3);
			END_FOR
		3:	// B3 bit through UNION + EXTENDS
			FOR k := 1 TO nIter DO
				GVL_Bench.dwSink := GVL_Bench.dwSink + BOOL_TO_DWORD(GVL_Bench.uExt.bits.bit3);
			END_FOR
		4:	// B4 bit through UNION
			FOR k := 1 TO nIter DO
				GVL_Bench.dwSink := GVL_Bench.dwSink + BOOL_TO_DWORD(GVL_Bench.uBits.bits.bit3);
			END_FOR
		5:	// B5 bit access to a WORD by dot
			FOR k := 1 TO nIter DO
				GVL_Bench.dwSink := GVL_Bench.dwSink + BOOL_TO_DWORD(GVL_Bench.wData.3);
			END_FOR
		6:	// B6 mask with a variable index
			FOR k := 1 TO nIter DO
				GVL_Bench.dwSink := GVL_Bench.dwSink + (SHR(GVL_Bench.dwDataB6, k AND 7) AND 1);
			END_FOR
		7:	// B7a: read 8 BOOL one after another (8 accesses per iteration)
			FOR k := 1 TO nIter DO
				GVL_Bench.dwSink := GVL_Bench.dwSink
					+ BOOL_TO_DWORD(GVL_Bench.stBools.b0) + BOOL_TO_DWORD(GVL_Bench.stBools.b1)
					+ BOOL_TO_DWORD(GVL_Bench.stBools.b2) + BOOL_TO_DWORD(GVL_Bench.stBools.b3)
					+ BOOL_TO_DWORD(GVL_Bench.stBools.b4) + BOOL_TO_DWORD(GVL_Bench.stBools.b5)
					+ BOOL_TO_DWORD(GVL_Bench.stBools.b6) + BOOL_TO_DWORD(GVL_Bench.stBools.b7);
			END_FOR
		8:	// B7b: read all 8 bits as one byte
			FOR k := 1 TO nIter DO
				GVL_Bench.dwSink := GVL_Bench.dwSink + BYTE_TO_DWORD(GVL_Bench.uBits.b);
			END_FOR
		9:	// B7c: read all 16 bits as one word
			FOR k := 1 TO nIter DO
				GVL_Bench.dwSink := GVL_Bench.dwSink + WORD_TO_DWORD(GVL_Bench.wData);
			END_FOR
		10:	// B8 bit of a WORD at an unaligned offset (pack_mode 0)
			FOR k := 1 TO nIter DO
				GVL_Bench.dwSink := GVL_Bench.dwSink + BOOL_TO_DWORD(GVL_Bench.stPacked.wData.3);
			END_FOR
		ELSE
			GVL_Bench.dwSink := GVL_Bench.dwSink + 1;
		END_CASE
	ELSE					// ---------- WRITE ----------
		CASE nVariant OF
		0:	// B0 baseline (the same shape as the write base)
			FOR k := 1 TO nIter DO
				GVL_Bench.dwSinkW := UDINT_TO_DWORD(k AND 1);
			END_FOR
		1:	// B1 BOOL field of a STRUCT
			FOR k := 1 TO nIter DO
				GVL_Bench.stBools.b3 := (k AND 1) <> 0;
			END_FOR
		2:	// B2 BIT field of a STRUCT
			FOR k := 1 TO nIter DO
				GVL_Bench.stBits.bit3 := (k AND 1) <> 0;
			END_FOR
		3:	// B3 bit through UNION + EXTENDS
			FOR k := 1 TO nIter DO
				GVL_Bench.uExt.bits.bit3 := (k AND 1) <> 0;
			END_FOR
		4:	// B4 bit through UNION
			FOR k := 1 TO nIter DO
				GVL_Bench.uBits.bits.bit3 := (k AND 1) <> 0;
			END_FOR
		5:	// B5 bit access to a WORD by dot
			FOR k := 1 TO nIter DO
				GVL_Bench.wData.3 := (k AND 1) <> 0;
			END_FOR
		6:	// B6 mask with a variable index (clear and set the bit)
			FOR k := 1 TO nIter DO
				GVL_Bench.dwDataB6 := (GVL_Bench.dwDataB6 AND NOT SHL(DWORD#1, k AND 7))
					OR SHL(BOOL_TO_DWORD((k AND 1) <> 0), k AND 7);
			END_FOR
		7:	// B7a group reset of 8 BOOL. The value depends on the previous one,
			// otherwise the compiler hoists the constant write out of the loop.
			FOR k := 1 TO nIter DO
				GVL_Bench.stBools.b0 := NOT GVL_Bench.stBools.b0;
				GVL_Bench.stBools.b1 := NOT GVL_Bench.stBools.b1;
				GVL_Bench.stBools.b2 := NOT GVL_Bench.stBools.b2;
				GVL_Bench.stBools.b3 := NOT GVL_Bench.stBools.b3;
				GVL_Bench.stBools.b4 := NOT GVL_Bench.stBools.b4;
				GVL_Bench.stBools.b5 := NOT GVL_Bench.stBools.b5;
				GVL_Bench.stBools.b6 := NOT GVL_Bench.stBools.b6;
				GVL_Bench.stBools.b7 := NOT GVL_Bench.stBools.b7;
			END_FOR
		8:	// B7b write all 8 bits as one byte (for the same reason - XOR)
			FOR k := 1 TO nIter DO
				GVL_Bench.uBits.b := GVL_Bench.uBits.b XOR BYTE#1;
			END_FOR
		9:	// B7c write all 16 bits as one word
			FOR k := 1 TO nIter DO
				GVL_Bench.wData := GVL_Bench.wData XOR WORD#1;
			END_FOR
		10:	// B8 write of a WORD bit at an unaligned offset (pack_mode 0)
			FOR k := 1 TO nIter DO
				GVL_Bench.stPacked.wData.3 := (k AND 1) <> 0;
			END_FOR
		ELSE
			GVL_Bench.dwSinkW := UDINT_TO_DWORD(k AND 1);
		END_CASE
	END_IF
END_IF

dwRes := SysTimeGetNs(t1);
tDur := t1 - t0;

END_FUNCTION_BLOCK

// PLC_Stabur/Application/F_Scale
FUNCTION F_Scale : REAL
VAR_INPUT
	x : REAL;
	k : REAL;
END_VAR

F_Scale := x * k;

END_FUNCTION

// PLC_Stabur/Application/FB_Logger
FUNCTION_BLOCK FB_Logger
VAR_INPUT
END_VAR
VAR_OUTPUT
END_VAR
VAR
	udiCmpId : UDINT;
	cmResult : Component_Manager.SysTypes.RTS_IEC_RESULT;
END_VAR

// Logger modelled on a production sample.
// Component registration and writing live in the methods LogADD / LogADDLong,
// so that the component name arrives as a parameter on every call.
// Log file on the PLC: /var/volatile/log/codesyscontrol.log

(*
Like LogADD, but for long strings: it cuts Message into pieces no longer than
CHUNK characters and writes each piece as a separate log record.
The runtime cuts a LogAdd2 record at 127 characters, hence CHUNK = 120.

The cut uses the built-in LEFT/RIGHT: copying characters one by one
(Short_Msg[i] := ...) does not advance the string length in CODESYS, and LogAdd2
receives an empty string - that is how the empty log records were produced.
*)

// LOG-file path: /var/volatile/log/codesyscontrol.log

METHOD LogADDLong : BOOL
VAR_INPUT
	Component : STRING;
	LogClass  : UDINT;
	Message   : STRING(1000) := 'something happened';
END_VAR
VAR CONSTANT
	CHUNK : INT := 120;		// chunk length, characters
END_VAR
VAR
	nLen  : INT;
	sRest : STRING(1000);
	sPart : STRING(255);
END_VAR
Component_Manager.CMAddComponent2(Component, 16#01, ADR(udiCmpId), ADR(cmResult));

sRest := Message;
nLen := LEN(sRest);

WHILE nLen > CHUNK DO
	sPart := LEFT(sRest, CHUNK);
	CmpLog.LogAdd2(cmplog.LogConstants.STD_LOGGER, udiCmpID, LogClass, cmpErrors.Errors.ERR_FAILED, 0, sPart);
	sRest := RIGHT(sRest, nLen - CHUNK);
	nLen := nLen - CHUNK;
END_WHILE

IF nLen > 0 THEN
	sPart := LEFT(sRest, nLen);
	CmpLog.LogAdd2(cmplog.LogConstants.STD_LOGGER, udiCmpID, LogClass, cmpErrors.Errors.ERR_FAILED, 0, sPart);
END_IF

LogADDLong := TRUE;
END_METHOD

(*
Like LogADD, but it watches the length itself: a string no longer than LIMIT
characters goes as one record, a longer one goes through LogADDLong in pieces.
The runtime cuts a LogAdd2 record at 127 characters, hence LIMIT = 120.
*)

// LOG-file path: /var/volatile/log/codesyscontrol.log

METHOD LogSafe : BOOL
VAR_INPUT
	Component : STRING;
	LogClass  : UDINT;
	Message   : STRING(255) := 'something happened';
END_VAR
VAR CONSTANT
	MAXLINE : INT := 120;	// LIMIT is an IEC reserved word, hence MAXLINE
END_VAR
IF LEN(Message) > MAXLINE THEN
	LogSafe := LogADDLong(Component, LogClass, Message);
ELSE
	LogSafe := LogADD(Component, LogClass, Message);
END_IF
END_METHOD

(*
Add new record in logfile
Component: STRING from LogComponent. Example: Component := LogComponent.BITBENCH
LogClass: CmpLog.LogClass. Example: LogClass := CmpLog.LogClass.LOG_ERROR
Message: STRING. Write here your Log Message.
*)

// LOG-file path: /var/volatile/log/codesyscontrol.log

METHOD LogADD : BOOL
VAR_INPUT
	Component : STRING;
	LogClass  : UDINT;
	Message   : STRING(255) := 'something happened';
END_VAR
Component_Manager.CMAddComponent2(Component, 16#01, ADR(udiCmpId), ADR(cmResult));

CmpLog.LogAdd2(cmplog.LogConstants.STD_LOGGER, udiCmpID, LogClass, cmpErrors.Errors.ERR_FAILED, 0, Message);
END_METHOD

(*
Prints an integer given in HUNDREDTHS (for example ns/operation * 100) as a
string with two places after the point: 1234 -> 12.34, -5 -> -0.05.
The result goes into LogComponent.sNumFmt: the call always has one argument.
*)

METHOD Fmt100 : BOOL
VAR_INPUT
	v		: DINT;
	xPlus	: BOOL := FALSE;	// TRUE: print positive values with a '+' sign
END_VAR
VAR
	xNeg    : BOOL;
	dwAbs   : DWORD;
	sBuf    : STRING(80);
	dwWhole : DWORD;
	dwFrac  : DWORD;
END_VAR
IF v < 0 THEN
	xNeg := TRUE;
	dwAbs := DINT_TO_DWORD(-v);
ELSE
	xNeg := FALSE;
	dwAbs := DINT_TO_DWORD(v);
END_IF

dwWhole := dwAbs / 100;
dwFrac  := dwAbs MOD 100;

sBuf := DWORD_TO_STRING(dwWhole);
sBuf := CONCAT(sBuf, '.');
IF dwFrac < 10 THEN
	sBuf := CONCAT(sBuf, '0');
END_IF
sBuf := CONCAT(sBuf, DWORD_TO_STRING(dwFrac));

IF xNeg THEN
	LogComponent.sNumFmt := CONCAT('-', sBuf);
ELSIF xPlus AND (v > 0) THEN
	LogComponent.sNumFmt := CONCAT('+', sBuf);
ELSE
	LogComponent.sNumFmt := sBuf;
END_IF

Fmt100 := TRUE;
END_METHOD

END_FUNCTION_BLOCK

// PLC_Stabur/Application/FB_Motor
FUNCTION_BLOCK FB_Motor
VAR_INPUT
	xStart : BOOL;
	xStop : BOOL;
	xFeedback : BOOL;
	xReset : BOOL;
	tFbTimeout : TIME := T#3S;
END_VAR
VAR_OUTPUT
	xRun : BOOL;
	xFault : BOOL;
	nStarts : UDINT;
END_VAR
VAR
	xStartPrev : BOOL;
	xResetPrev : BOOL;
	xStartRise : BOOL;
	xResetRise : BOOL;
	xAwaitingFeedback : BOOL;
	tFeedback : TON;
END_VAR

xStartRise := xStart AND NOT xStartPrev;
xResetRise := xReset AND NOT xResetPrev;
xStartPrev := xStart;
xResetPrev := xReset;

tFeedback(IN := xAwaitingFeedback, PT := tFbTimeout);

IF xResetRise THEN
	xFault := FALSE;
	xRun := FALSE;
	xAwaitingFeedback := FALSE;
END_IF

IF xStop THEN
	xRun := FALSE;
	xAwaitingFeedback := FALSE;
ELSIF xFault THEN
	xRun := FALSE;
	xAwaitingFeedback := FALSE;
ELSIF xRun AND NOT xAwaitingFeedback THEN
	IF NOT xFeedback THEN
		xRun := FALSE;
		xFault := TRUE;
	END_IF
ELSIF xAwaitingFeedback THEN
	IF tFeedback.Q THEN
		xRun := FALSE;
		xAwaitingFeedback := FALSE;
		xFault := TRUE;
	ELSIF xFeedback THEN
		xAwaitingFeedback := FALSE;
		nStarts := nStarts + 1;
	END_IF
ELSIF xStartRise THEN
	xRun := TRUE;
	xAwaitingFeedback := TRUE;
END_IF

END_FUNCTION_BLOCK

// PLC_Stabur/Application/FB_Valve
FUNCTION_BLOCK FB_Valve
VAR
	xOpen : BOOL;
END_VAR

PROPERTY P_Open : BOOL
GET
P_Open := xOpen;
END_GET
SET
xOpen := P_Open;
END_SET
END_PROPERTY

ACTION A_Reset:
xOpen := FALSE;
END_ACTION

METHOD M_Toggle : BOOL
xOpen := NOT xOpen;
M_Toggle := xOpen;
END_METHOD

END_FUNCTION_BLOCK

// PLC_Stabur/Application/I_LiveTmp
INTERFACE I_LiveTmp

METHOD M_LiveTmp : BOOL
VAR_INPUT
	x : BOOL;
END_VAR
END_METHOD

END_INTERFACE

// PLC_Stabur/Application/Visualization
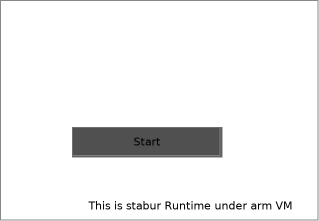
VISUALIZATION Visualization  // 319x221
    Button (72,127 150x30), "Start"
    Label (62,191 257x30), "This is stabur Runtime under arm VM"
END_VISUALIZATION
